// Einzige Schnittstelle des Ablaufs zur Achskopplung. Details: docs/kinematik.md
INTERFACE I_Kinematics

METHOD Cyclic
// Einmal pro SPS-Zyklus aufrufen.
VAR_INPUT
END_VAR
END_METHOD

METHOD LoadPlan : BOOL
// Aktiven Plan (GVL_Plan.stActive) mit dieser ID übernehmen. Nur entkoppelt.
VAR_INPUT
    nPlanId : UDINT;
END_VAR
END_METHOD

METHOD LoadSection : BOOL
// Kurvenscheiben des Abschnitts nSection laden. Nur entkoppelt; fertig, wenn TableReady() TRUE meldet.
VAR_INPUT
    nSection : INT;
END_VAR
END_METHOD

METHOD TableReady : BOOL
VAR_INPUT
END_VAR
END_METHOD

METHOD Start : BOOL
// Koppelt X und A an Z1 und startet den Master.
VAR_INPUT
END_VAR
END_METHOD

METHOD Hold : BOOL
// Bremst den Master. Die Kopplung bleibt bestehen.
VAR_INPUT
END_VAR
END_METHOD

METHOD Resume : BOOL
// Setzt den Master aus dem Halt fort (nicht an einer offenen Rotation oder am Abschnittsende).
VAR_INPUT
END_VAR
END_METHOD

METHOD AtRotation : BOOL
// Master steht an einer Rotationsposition; RotationAngle() liefert den Drehwinkel für W.
VAR_INPUT
END_VAR
END_METHOD

METHOD RotationAngle : LREAL
VAR_INPUT
END_VAR
END_METHOD

METHOD ContinueAfterRotation : BOOL
VAR_INPUT
END_VAR
END_METHOD

METHOD SectionDone : BOOL
// Master steht am Ende des Abschnitts, Kopplung besteht noch.
VAR_INPUT
END_VAR
END_METHOD

METHOD Abort : BOOL
// Stoppt den Master und löst die Kopplung.
VAR_INPUT
END_VAR
END_METHOD

METHOD Reset : BOOL
// Quittiert einen Fehler der Kinematik. Der Plan bleibt erhalten.
VAR_INPUT
END_VAR
END_METHOD

METHOD Unload : BOOL
// Plan verwerfen (nur entkoppelt).
VAR_INPUT
END_VAR
END_METHOD

METHOD IsCoupled : BOOL
VAR_INPUT
END_VAR
END_METHOD

METHOD GetStatus : ST_KinStatus
VAR_INPUT
END_VAR
END_METHOD

END_INTERFACE

(* stored: Version 1.1.0.1
   Itf I_Kinematics: Id {c5693eee-b791-4378-8103-14055035bf96}
   Method Cyclic: Id {5ff6501c-e7b5-5368-a3a5-5426dfc9aa2c}
   Method LoadPlan: Id {a7d084e2-8bb5-5cd6-ab5b-bbfad6b21f43}
   Method LoadSection: Id {3dfa17f9-91ed-5fc6-8a1a-bd2b1ac01ae8}
   Method TableReady: Id {d8fceddd-56a1-5270-932b-97cdf7569951}
   Method Start: Id {d830ff77-cb65-5116-9c0a-2bfdcec02fd3}
   Method Hold: Id {96cda0db-d84f-5c41-8a73-c4e3bd3aa973}
   Method Resume: Id {6d8827b9-0e6a-5f1e-a3c5-9876d793655f}
   Method AtRotation: Id {460217e9-8a87-5886-918f-8533ac6f4f8c}
   Method RotationAngle: Id {f76901e6-6a2f-55de-a766-78d83766bfe6}
   Method ContinueAfterRotation: Id {b7699b80-92df-5aad-8221-cd28c18d69e8}
   Method SectionDone: Id {9ee8b7a2-2774-5239-8ca5-ea486bb079d4}
   Method Abort: Id {c807c0fd-8651-58b7-800f-706843c63d1b}
   Method Reset: Id {98e116bc-6e51-5ba3-88fe-239e21efc8ff}
   Method Unload: Id {ee67441f-f2dd-5594-a8a8-d045785b30b4}
   Method IsCoupled: Id {9fe684e1-fcf7-513c-8ee7-b2d21522eeb3}
   Method GetStatus: Id {01362359-882e-5793-8949-44ea05380c9a} *)
